FUNCTION_BLOCK AOption_X_TO_EVENT (* Composite FB for convert AOption to EVENT (Fan-In, haelt den SOCKET) *)
  (* Standard: 61499-2; Description: Copyright (c) 2026 Meisterschulen am Ostbahnhof This program and the accompanying materials are made available under the terms of the Eclipse Public License 2.0 which is available at https://www.eclipse.org/legal/epl-2.0/ SPDX-License-Identifier: EPL-2.0 *)
  (* Version 1.0, 2026-10-13, Franz Höpfinger, Meisterschulen am Ostbahnhof *)
  PACKAGE Option::conversion;
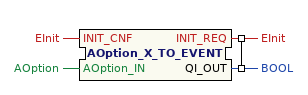
  EVENT_INPUT
    INIT_CNF : EInit; (* Confirmation to Adapter *)
  END_EVENT
  EVENT_OUTPUT
    INIT_REQ : EInit WITH QI_OUT; (* Request from Adapter *)
  END_EVENT
  VAR_OUTPUT
    QI_OUT : BOOL; (* Event Input Qualifier (IEC 61499-1): TRUE=Option anfordern/aktivieren, FALSE=zurueckziehen *)
  END_VAR
  SOCKETS
    AOption_IN : Option::AOption; (* Adapter Input *)
  END_SOCKETS
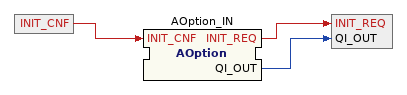
  EVENT_CONNECTIONS
    AOption_IN.INIT_REQ TO INIT_REQ;
    INIT_CNF TO AOption_IN.INIT_CNF;
  END_CONNECTIONS
  DATA_CONNECTIONS
    AOption_IN.QI_OUT TO QI_OUT;
  END_CONNECTIONS
END_FUNCTION_BLOCK
